(* IEC 61131-3 sources: Test-Git_ESME26/TestProgettoESME_26.fbsproj/PacDriveLib Migration/Motion/Homing/PDL_FB_ResetTrackingDeviation.fb.st^, 3 files *)

(* ---- ifDrive2.prop.st ---- *)
PROPERTY PUBLIC ifDrive2 : DDI.IF_Drive2;

__SETTERDECLARATION__
VAR
END_VAR
__SETTERIMPLEMENTATION__
ifDrive2_loc := ifDrive2;

(* ---- lrOldTrackDevLim.prop.st ---- *)
PROPERTY PUBLIC lrOldTrackDevLim : LREAL
__SETTERDECLARATION__
VAR
END_VAR
__SETTERIMPLEMENTATION__
lrOldTrackingDeviationLimit := lrOldTrackDevLim;
__GETTERDECLARATION__
VAR
END_VAR
__GETTERIMPLEMENTATION__

(* ---- xDone.prop.st ---- *)
PROPERTY xDone : BOOL
__GETTERDECLARATION__
VAR
END_VAR
__GETTERIMPLEMENTATION__
xDone := xDone_loc;
__SETTERDECLARATION__
VAR
END_VAR
__SETTERIMPLEMENTATION__
xDone_loc := xDone;
